{attribute 'linkalways'} 
{attribute 'no_explicit_call' := 'This FB is a CLASS and must be accessed using methods or properties'}
{attribute 'enable_dynamic_creation'}
FUNCTION_BLOCK _ETcVnNormalizationType EXTENDS EnumDatatypeBase
VAR
	localData : ETcVnNormalizationType;
	activeData : REFERENCE TO ETcVnNormalizationType;
	enumBaseDatatype : _DINT(localData);
END_VAR

METHOD PRIVATE AddLocalEnumeration
VAR_INPUT
	Enumeration : T_MAXSTRING;
	Value : ETcVnNormalizationType;
END_VAR
AddEnumeration(Enumeration, Value);
END_METHOD

PROPERTY PUBLIC Address : PVOID
GET
Address := ADR(activeData);
END_GET
END_PROPERTY

METHOD PUBLIC ClearReference
VAR_INPUT
END_VAR
activeData REF= localData;
SetBaseDatatypeReference();
END_METHOD

METHOD PUBLIC Clone : I_Datatype
VAR
    pClone : POINTER TO _ETcVnNormalizationType;
END_VAR
pClone := __NEW(_ETcVnNormalizationType(InitialValue := Value));
Clone := pClone^;
END_METHOD

METHOD FB_init : BOOL
VAR_INPUT
	bInitRetains : BOOL; // if TRUE, the retain variables are initialized (warm start / cold start)
	bInCopyCode : BOOL;  // if TRUE, the instance afterwards gets moved into the copy code (online change)
	InitialValue : ETcVnNormalizationType;
END_VAR
localData := InitialValue;
AddBaseDatatype(enumBaseDatatype);
ClearReference();

AddLocalEnumeration('TCVN_NT_INF', ETcVnNormalizationType.TCVN_NT_INF);
AddLocalEnumeration('TCVN_NT_L1', ETcVnNormalizationType.TCVN_NT_L1);
AddLocalEnumeration('TCVN_NT_L2', ETcVnNormalizationType.TCVN_NT_L2);
AddLocalEnumeration('TCVN_NT_L2SQR', ETcVnNormalizationType.TCVN_NT_L2SQR);
AddLocalEnumeration('TCVN_NT_HAMMING', ETcVnNormalizationType.TCVN_NT_HAMMING);
AddLocalEnumeration('TCVN_NT_HAMMING2', ETcVnNormalizationType.TCVN_NT_HAMMING2);
AddLocalEnumeration('TCVN_NT_RELATIVE_INF', ETcVnNormalizationType.TCVN_NT_RELATIVE_INF);
AddLocalEnumeration('TCVN_NT_RELATIVE_L1', ETcVnNormalizationType.TCVN_NT_RELATIVE_L1);
AddLocalEnumeration('TCVN_NT_RELATIVE_L2', ETcVnNormalizationType.TCVN_NT_RELATIVE_L2);
AddLocalEnumeration('TCVN_NT_RELATIVE_L2SQR', ETcVnNormalizationType.TCVN_NT_RELATIVE_L2SQR);
AddLocalEnumeration('TCVN_NT_RELATIVE_HAMMING', ETcVnNormalizationType.TCVN_NT_RELATIVE_HAMMING);
AddLocalEnumeration('TCVN_NT_RELATIVE_HAMMING2', ETcVnNormalizationType.TCVN_NT_RELATIVE_HAMMING2);
AddLocalEnumeration('TCVN_NT_MINMAX', ETcVnNormalizationType.TCVN_NT_MINMAX);
END_METHOD

PROPERTY PUBLIC Identifier : T_MAXSTRING
GET
Identifier := 'ETcVnNormalizationType';
END_GET
END_PROPERTY

METHOD IsEnumeratorValueEqual : BOOL
VAR_INPUT
	Enumerator : I_KeyValueForwardEnumerator;
END_VAR
VAR
	storedValue : ETcVnNormalizationType;
END_VAR
IF NOT Enumerator.TryGet(storedValue) THEN
	RETURN;
END_IF

IsEnumeratorValueEqual := storedValue = activeData;
END_METHOD

METHOD PUBLIC MakeReferenceTo
VAR_INPUT
	ReferenceTarget : REFERENCE TO ETcVnNormalizationType;
END_VAR
activeData REF= ReferenceTarget;
SetBaseDatatypeReference();
END_METHOD

METHOD PROTECTED SetBaseDatatypeReference
VAR_INPUT
END_VAR
enumBaseDatatype.MakeReferenceTo(activeData);
END_METHOD

PROPERTY PUBLIC Size : UDINT
GET
Size := SIZEOF(activeData);
END_GET
END_PROPERTY

METHOD TryMakeReferenceTo : BOOL
VAR_INPUT
	Target : I_Datatype;
END_VAR
VAR
	pTargetData : POINTER TO ETcVnNormalizationType;
END_VAR
IF NOT IsEquivalentTo(Target) THEN
	RETURN;
END_IF

pTargetData := Target.Address;
activeData REF= pTargetData^;
SetBaseDatatypeReference();
TryMakeReferenceTo := TRUE;
END_METHOD

PROPERTY PUBLIC Value : ETcVnNormalizationType
GET
Value := activeData;
END_GET
SET
activeData := Value;
END_SET
END_PROPERTY

END_FUNCTION_BLOCK

(* stored: Version 1.1.0.1, ProductVersion 3.1.4024.13
   POU _ETcVnNormalizationType: Id {091b2290-906a-0fa8-2950-956d64c3c8f0}, SpecialFunc None
   Folder Core: Id {00df3bb2-6758-026f-360a-5723cc35778f}
   Folder Protected: Id {37deeed4-0c25-0f3b-2ccb-4b50385dd6ae}
   Folder Customize: Id {2208d4a6-2f2a-0b15-2472-63f6d552d68b}
   Folder Constructor: Id {eb5bb077-1ce4-0e9b-34ec-141f24370e6d}
   Folder Private: Id {43cc0a02-36f0-05fe-284f-8866b2243e46}
   Folder Protected: Id {294dc737-79ec-0e54-3bcb-795e978dab90}
   Method AddLocalEnumeration: Id {0bd783e2-4a72-072d-0c59-bb359da507f8}
   Property Address: Id {b9c34c68-d0b7-0e5b-034e-3efc3203b069}
   Get Get: Id {2490cce1-adf3-0b96-2d3a-1db67fa6f832}
   Method ClearReference: Id {d5ca2dc2-3f9f-0b48-2149-34f95734db1f}
   Method Clone: Id {1b921516-b9cf-0831-262b-0d83d9e2a536}
   Method FB_init: Id {daedd4da-5a57-0008-0325-220534e4d3e0}
   Property Identifier: Id {4f7deeb6-aa29-0df6-338f-7a0d50a0f78b}
   Get Get: Id {218c77a5-5bfd-06f9-122b-daa34d9c536f}
   Method IsEnumeratorValueEqual: Id {9f7b3d8b-fcd7-0735-3842-783ed62a7ff0}
   Method MakeReferenceTo: Id {1853454e-5161-01ff-2de5-e27abaaae5bf}
   Method SetBaseDatatypeReference: Id {57485417-756d-0a92-0061-439256603162}
   Property Size: Id {dce8127b-27e7-0532-25e3-6d0c1f150326}
   Get Get: Id {c3267c9c-dbc4-08c8-1eba-8f377440d0a4}
   Method TryMakeReferenceTo: Id {f10ffc1f-c49f-0bad-1875-911122058f9d}
   Property Value: Id {0249c051-cdd0-02fd-2100-206c2fa70cd3}
   Get Get: Id {431c27d1-9b7c-0621-1cf9-a48cb71a829a}
   Set Set: Id {11831029-b79d-0847-24f6-90151c36089e} *)
